// TIA Portal V21 export
// export: Created 2026-11-10T19:11:33.3480051Z, ExportSetting WithDefaults, DisplayName Totally Integrated Automation Portal, DisplayVersion V21 Update 3, DisplayName STEP 7 Professional, DisplayVersion V21 Update 3, DisplayName STEP 7 Safety, DisplayVersion V21, DisplayName Tech WebApplication, DisplayVersion V21, DisplayName WinCC Basic/Comfort/Advanced, DisplayVersion V21 Update 3, DisplayName WinCC Unified, DisplayVersion V21 Update 3
DATA_BLOCK "DB_TRCV_C"   // DB10
// stored: AutoNumber true, DBAccessibleFromOPCUA true, DBAccessibleFromWebserver true, InstanceOfName TRCV_C, OfSystemLibElement TRCV_C, OfSystemLibVersion 3.2
"TRCV_C"
   // VAR_INPUT
   //    EN_R : Bool;
   //    CONT : Bool;
   //    LEN : UDInt;
   //    ADHOC : Bool;
   // END_VAR
   // VAR_OUTPUT
   //    DONE : Bool;
   //    BUSY : Bool;
   //    ERROR : Bool;
   //    STATUS : Word;
   //    RCVD_LEN : UDInt;
   // END_VAR
   // VAR_IN_OUT
   //    CONNECT : Variant;
   //    DATA : Variant;
   //    ADDR : Variant;
   //    COM_RST : Bool;
   // END_VAR
   // VAR
   //    s_state : Int;
   //    s_locked : Bool;
   //    s_udp : Bool;
   //    s_configured : Bool;
   //    s_tcon_80A3 : Bool;
   //    s_ConID : CONN_OUC;
   //    s_TCON { S7_SetPoint := 'True'} : TCON;
   //    s_TDIAG { S7_SetPoint := 'True'} : T_DIAG;
   //    s_TDIAG_Status { S7_SetPoint := 'True'} : TDiag_Status;
   //    s_TRCV { S7_SetPoint := 'True'} : TRCV;
   //    s_TURCV { S7_SetPoint := 'True'} : TURCV;
   //    s_TDISCON { S7_SetPoint := 'True'} : TDISCON;
   //    s_TRESET { S7_SetPoint := 'True'} : T_RESET;
   // END_VAR
BEGIN
END_DATA_BLOCK
